{attribute 'qualified_only'}
{attribute 'strict'}
{attribute 'to_string'}
TYPE E_FileExporterState :
(
	error := -10,
	idle := 0,
	serializing := 10,
	creating := 15,
	opening := 20,
	buffering := 25,
	writing := 30,
	closing := 40,
	rotating := 50,
	done := 99
);
END_TYPE
//  error = '-10'

(* stored: Version 1.1.0.1
   EnumerationTextList E_FileExporterState: Id {f847849e-dedd-4c0a-8d83-974df81b7fcb} *)
